Staubli VAL3: start.pgx

program start()
begin
  call home:main()
end
